// TIA Portal V21 export
// export: Created 2026-11-07T14:35:58.367327Z, ExportSetting WithDefaults, DisplayName Totally Integrated Automation Portal, DisplayVersion V21, DisplayName STEP 7 Professional, DisplayVersion V21, DisplayName STEP 7 Safety, DisplayVersion V21, DisplayName Tech WebApplication, DisplayVersion V21, DisplayName WinCC Basic/Comfort/Advanced, DisplayVersion V21, DisplayName WinCC Unified, DisplayVersion V21
Screen "T01_Rect"  1024x768, Number=21
  ScreenLayer 
    Rectangle "P_CellRect" at 0,0 size 100x30  StyleItem=Rectangle
